(* PLC project GeneratedProgram, SafePLC-Gen SafePLC-Gen Multimodal 1.0 *)
(* stored: creationDateTime 2026-04-25T13:21:32.531016Z *)

PROGRAM GeneratedProgram
  VAR
    PI_4712_01_Scaled : REAL;
    PICSA_4712_02_Scaled : REAL;
    TICSA_4750_03_Scaled : REAL;
    PI_4712_01_EU_Min : REAL;
    PI_4712_01_EU_Span : REAL;
    PICSA_4712_02_EU_Min : REAL;
    PICSA_4712_02_EU_Span : REAL;
    TICSA_4750_03_EU_Min : REAL;
    TICSA_4750_03_EU_Span : REAL;
    PI_4712_01_HH_SP : REAL;
    PI_4712_01_H_SP : REAL;
    PI_4712_01_L_SP : REAL;
    PI_4712_01_LL_SP : REAL;
    PI_4712_01_Deadband : REAL;
    PI_4712_01_HH : BOOL;
    PI_4712_01_H : BOOL;
    PI_4712_01_L : BOOL;
    PI_4712_01_LL : BOOL;
    PI_4712_01_HH_Latch : SR;
    PI_4712_01_LL_Latch : SR;
    PI_4712_01_HH_Ack : BOOL;
    PI_4712_01_LL_Ack : BOOL;
    PICSA_4712_02_HH_SP : REAL;
    PICSA_4712_02_H_SP : REAL;
    PICSA_4712_02_L_SP : REAL;
    PICSA_4712_02_LL_SP : REAL;
    PICSA_4712_02_Deadband : REAL;
    PICSA_4712_02_HH : BOOL;
    PICSA_4712_02_H : BOOL;
    PICSA_4712_02_L : BOOL;
    PICSA_4712_02_LL : BOOL;
    PICSA_4712_02_HH_Latch : SR;
    PICSA_4712_02_LL_Latch : SR;
    PICSA_4712_02_HH_Ack : BOOL;
    PICSA_4712_02_LL_Ack : BOOL;
    PICSA_4712_02_SP : REAL;
    PICSA_4712_02_Kp : REAL;
    PICSA_4712_02_Ki : REAL;
    PICSA_4712_02_Error : REAL;
    PICSA_4712_02_Integ : REAL;
    PICSA_4712_02_Output : REAL;
    TICSA_4750_03_HH_SP : REAL;
    TICSA_4750_03_H_SP : REAL;
    TICSA_4750_03_L_SP : REAL;
    TICSA_4750_03_LL_SP : REAL;
    TICSA_4750_03_Deadband : REAL;
    TICSA_4750_03_HH : BOOL;
    TICSA_4750_03_H : BOOL;
    TICSA_4750_03_L : BOOL;
    TICSA_4750_03_LL : BOOL;
    TICSA_4750_03_HH_Latch : SR;
    TICSA_4750_03_LL_Latch : SR;
    TICSA_4750_03_HH_Ack : BOOL;
    TICSA_4750_03_LL_Ack : BOOL;
    TICSA_4750_03_SP : REAL;
    TICSA_4750_03_Kp : REAL;
    TICSA_4750_03_Ki : REAL;
    TICSA_4750_03_Error : REAL;
    TICSA_4750_03_Integ : REAL;
    TICSA_4750_03_Output : REAL;
    HV4750_01_Out : BOOL;
    System_Alarm : BOOL;
    FirstScan : BOOL;
  END_VAR

            IF FirstScan THEN
    PV4712_02_Out        := 6554;
    TV4750_03_Out        := 6554;
    HV4750_01_Out        := FALSE;
    PICSA_4712_02_Integ  := 0.0;
    TICSA_4750_03_Integ  := 0.0;
    PI_4712_01_HH_Latch(S1 := FALSE, R := FALSE);
    PI_4712_01_LL_Latch(S1 := FALSE, R := FALSE);
    PICSA_4712_02_HH_Latch(S1 := FALSE, R := FALSE);
    PICSA_4712_02_LL_Latch(S1 := FALSE, R := FALSE);
    TICSA_4750_03_HH_Latch(S1 := FALSE, R := FALSE);
    TICSA_4750_03_LL_Latch(S1 := FALSE, R := FALSE);
    FirstScan            := FALSE;
    RETURN;
END_IF;

PI_4712_01_Scaled    := ((INT_TO_REAL(PI_4712_01_Raw)    - 6554.0) / (32767.0 - 6554.0)) * PI_4712_01_EU_Span    + PI_4712_01_EU_Min;
PICSA_4712_02_Scaled := ((INT_TO_REAL(PICSA_4712_02_Raw) - 6554.0) / (32767.0 - 6554.0)) * PICSA_4712_02_EU_Span + PICSA_4712_02_EU_Min;
TICSA_4750_03_Scaled := ((INT_TO_REAL(TICSA_4750_03_Raw) - 6554.0) / (32767.0 - 6554.0)) * TICSA_4750_03_EU_Span + TICSA_4750_03_EU_Min;

(* PI-4712.01 alarms — monitoring only *)
IF PI_4712_01_Scaled >= PI_4712_01_HH_SP THEN
    PI_4712_01_HH := TRUE;
    PI_4712_01_HH_Latch(S1 := TRUE, R := FALSE);
ELSIF PI_4712_01_Scaled <= (PI_4712_01_HH_SP - PI_4712_01_Deadband) THEN
    PI_4712_01_HH := FALSE;
    PI_4712_01_HH_Latch(S1 := FALSE, R := (PI_4712_01_HH_Ack AND NOT PI_4712_01_HH));
END_IF;

IF PI_4712_01_Scaled >= PI_4712_01_H_SP THEN
    PI_4712_01_H := TRUE;
ELSIF PI_4712_01_Scaled < (PI_4712_01_H_SP - PI_4712_01_Deadband) THEN
    PI_4712_01_H := FALSE;
END_IF;

IF PI_4712_01_Scaled <= PI_4712_01_L_SP THEN
    PI_4712_01_L := TRUE;
ELSIF PI_4712_01_Scaled > (PI_4712_01_L_SP + PI_4712_01_Deadband) THEN
    PI_4712_01_L := FALSE;
END_IF;

IF PI_4712_01_Scaled <= PI_4712_01_LL_SP THEN
    PI_4712_01_LL := TRUE;
    PI_4712_01_LL_Latch(S1 := TRUE, R := FALSE);
ELSIF PI_4712_01_Scaled >= (PI_4712_01_LL_SP + PI_4712_01_Deadband) THEN
    PI_4712_01_LL := FALSE;
    PI_4712_01_LL_Latch(S1 := FALSE, R := (PI_4712_01_LL_Ack AND NOT PI_4712_01_LL));
END_IF;

(* PICSA-4712.02 alarms *)
IF PICSA_4712_02_Scaled >= PICSA_4712_02_HH_SP THEN
    PICSA_4712_02_HH := TRUE;
    PICSA_4712_02_HH_Latch(S1 := TRUE, R := FALSE);
ELSIF PICSA_4712_02_Scaled <= (PICSA_4712_02_HH_SP - PICSA_4712_02_Deadband) THEN
    PICSA_4712_02_HH := FALSE;
    PICSA_4712_02_HH_Latch(S1 := FALSE, R := (PICSA_4712_02_HH_Ack AND NOT PICSA_4712_02_HH));
END_IF;

IF PICSA_4712_02_Scaled >= PICSA_4712_02_H_SP THEN
    PICSA_4712_02_H := TRUE;
ELSIF PICSA_4712_02_Scaled < (PICSA_4712_02_H_SP - PICSA_4712_02_Deadband) THEN
    PICSA_4712_02_H := FALSE;
END_IF;

IF PICSA_4712_02_Scaled <= PICSA_4712_02_L_SP THEN
    PICSA_4712_02_L := TRUE;
ELSIF PICSA_4712_02_Scaled > (PICSA_4712_02_L_SP + PICSA_4712_02_Deadband) THEN
    PICSA_4712_02_L := FALSE;
END_IF;

IF PICSA_4712_02_Scaled <= PICSA_4712_02_LL_SP THEN
    PICSA_4712_02_LL := TRUE;
    PICSA_4712_02_LL_Latch(S1 := TRUE, R := FALSE);
ELSIF PICSA_4712_02_Scaled >= (PICSA_4712_02_LL_SP + PICSA_4712_02_Deadband) THEN
    PICSA_4712_02_LL := FALSE;
    PICSA_4712_02_LL_Latch(S1 := FALSE, R := (PICSA_4712_02_LL_Ack AND NOT PICSA_4712_02_LL));
END_IF;

(* PICSA-4712.02 PI pressure controller → PV4712.02 *)
PICSA_4712_02_Error  := PICSA_4712_02_SP - PICSA_4712_02_Scaled;
PICSA_4712_02_Integ  := PICSA_4712_02_Integ + (PICSA_4712_02_Ki * PICSA_4712_02_Error);
IF PICSA_4712_02_Integ > 100.0 THEN
    PICSA_4712_02_Integ := 100.0;
ELSIF PICSA_4712_02_Integ < 0.0 THEN
    PICSA_4712_02_Integ := 0.0;
END_IF;
PICSA_4712_02_Output := (PICSA_4712_02_Kp * PICSA_4712_02_Error) + PICSA_4712_02_Integ;
IF PICSA_4712_02_Output > 100.0 THEN
    PICSA_4712_02_Output := 100.0;
ELSIF PICSA_4712_02_Output < 0.0 THEN
    PICSA_4712_02_Output := 0.0;
END_IF;
PV4712_02_Out := REAL_TO_INT(6554.0 + (PICSA_4712_02_Output / 100.0) * (32767.0 - 6554.0));

(* TICSA-4750.03 alarms *)
IF TICSA_4750_03_Scaled >= TICSA_4750_03_HH_SP THEN
    TICSA_4750_03_HH := TRUE;
    TICSA_4750_03_HH_Latch(S1 := TRUE, R := FALSE);
ELSIF TICSA_4750_03_Scaled <= (TICSA_4750_03_HH_SP - TICSA_4750_03_Deadband) THEN
    TICSA_4750_03_HH := FALSE;
    TICSA_4750_03_HH_Latch(S1 := FALSE, R := (TICSA_4750_03_HH_Ack AND NOT TICSA_4750_03_HH));
END_IF;

IF TICSA_4750_03_Scaled >= TICSA_4750_03_H_SP THEN
    TICSA_4750_03_H := TRUE;
ELSIF TICSA_4750_03_Scaled < (TICSA_4750_03_H_SP - TICSA_4750_03_Deadband) THEN
    TICSA_4750_03_H := FALSE;
END_IF;

IF TICSA_4750_03_Scaled <= TICSA_4750_03_L_SP THEN
    TICSA_4750_03_L := TRUE;
ELSIF TICSA_4750_03_Scaled > (TICSA_4750_03_L_SP + TICSA_4750_03_Deadband) THEN
    TICSA_4750_03_L := FALSE;
END_IF;

IF TICSA_4750_03_Scaled <= TICSA_4750_03_LL_SP THEN
    TICSA_4750_03_LL := TRUE;
    TICSA_4750_03_LL_Latch(S1 := TRUE, R := FALSE);
ELSIF TICSA_4750_03_Scaled >= (TICSA_4750_03_LL_SP + TICSA_4750_03_Deadband) THEN
    TICSA_4750_03_LL := FALSE;
    TICSA_4750_03_LL_Latch(S1 := FALSE, R := (TICSA_4750_03_LL_Ack AND NOT TICSA_4750_03_LL));
END_IF;

(* TICSA-4750.03 PI temperature controller → TV4750.03 *)
TICSA_4750_03_Error  := TICSA_4750_03_SP - TICSA_4750_03_Scaled;
TICSA_4750_03_Integ  := TICSA_4750_03_Integ + (TICSA_4750_03_Ki * TICSA_4750_03_Error);
IF TICSA_4750_03_Integ > 100.0 THEN
    TICSA_4750_03_Integ := 100.0;
ELSIF TICSA_4750_03_Integ < 0.0 THEN
    TICSA_4750_03_Integ := 0.0;
END_IF;
TICSA_4750_03_Output := (TICSA_4750_03_Kp * TICSA_4750_03_Error) + TICSA_4750_03_Integ;
IF TICSA_4750_03_Output > 100.0 THEN
    TICSA_4750_03_Output := 100.0;
ELSIF TICSA_4750_03_Output < 0.0 THEN
    TICSA_4750_03_Output := 0.0;
END_IF;
TV4750_03_Out := REAL_TO_INT(6554.0 + (TICSA_4750_03_Output / 100.0) * (32767.0 - 6554.0));

(* HS-4750.01 hand switch drives HV4750.01 directly *)
HV4750_01_Out := HS_4750_01;

(* Aggregate all alarm states — consumed by SCADA/HMI *)
System_Alarm :=
    PI_4712_01_HH_Latch.Q1 OR PI_4712_01_LL_Latch.Q1 OR
    PI_4712_01_H            OR PI_4712_01_L            OR
    PI_4712_01_HH           OR PI_4712_01_LL           OR
    PICSA_4712_02_HH_Latch.Q1 OR PICSA_4712_02_LL_Latch.Q1 OR
    PICSA_4712_02_H            OR PICSA_4712_02_L            OR
    PICSA_4712_02_HH           OR PICSA_4712_02_LL           OR
    TICSA_4750_03_HH_Latch.Q1 OR TICSA_4750_03_LL_Latch.Q1 OR
    TICSA_4750_03_H            OR TICSA_4750_03_L            OR
    TICSA_4750_03_HH           OR TICSA_4750_03_LL;
          
END_PROGRAM

CONFIGURATION Config0
  RESOURCE Res0 ON PLC
    TASK MainTask(INTERVAL := T#20ms, PRIORITY := 0);
    PROGRAM Main : GeneratedProgram;
  END_RESOURCE
END_CONFIGURATION
